SUBAPPLICATION Uebung_OPC_L16b_AX (* Wie L16, aber: gelesen wird erst, wenn INCREMENTED die Berechnung gemeldet hat (statt direkt nach dem Schreiben) *)
  (* Standard: 61499-2; Description: Copyright (c) 2026 Meisterschulen am Ostbahnhof This program and the accompanying materials are made available under the terms of the Eclipse Public License 2.0 which is available at https://www.eclipse.org/legal/epl-2.0/ SPDX-License-Identifier: EPL-2.0 *)
  (* Version 1.0, 2026-10-18, Franz Höpfinger, Meisterschulen am Ostbahnhof, B-Version von L16: Lesen erst nach INCREMENTED.CNF *)
  PACKAGE Meins::OPC_UA_Lokal;
  IMPORT Meins::OPC_UA_Lokal::const::OpcUaLokal::L16B_INC_READ;
  IMPORT Meins::OPC_UA_Lokal::const::OpcUaLokal::L16B_INCD_WRITE;
  IMPORT Meins::OPC_UA_Lokal::const::OpcUaLokal::L16B_INC_CLIENT_WRITE;
  IMPORT Meins::OPC_UA_Lokal::const::OpcUaLokal::L16B_INCD_CLIENT_READ;
  IMPORT logiBUS::io::DI::logiBUS_DI::Input_I1;
  IMPORT logiBUS::io::DI::logiBUS_DI_Events::BUTTON_PRESS_DOWN;
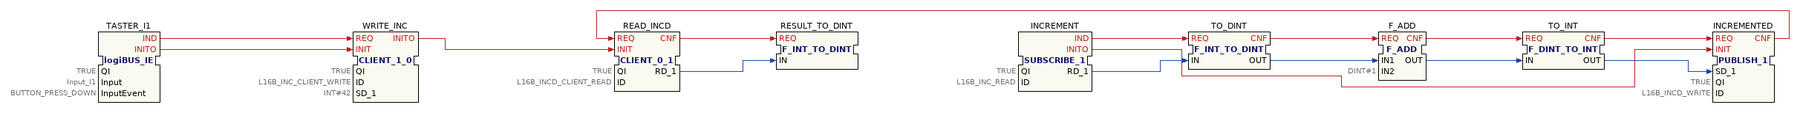
  (* B-Version von Uebung_OPC_L16_AX: READ_INCD.REQ kommt von INCREMENTED.CNF (Ergebnis ist veroeffentlicht), nicht von WRITE_INC.CNF. Das Lesen haengt so nicht mehr von der Reihenfolge ab. *)
  FBS
    TASTER_I1 : logiBUS::io::DI::logiBUS_IE(QI := TRUE, Input := Input_I1, InputEvent := BUTTON_PRESS_DOWN);
    WRITE_INC : iec61499::net::CLIENT_1_0(QI := TRUE, ID := L16B_INC_CLIENT_WRITE, SD_1 := INT#42);
    READ_INCD : iec61499::net::CLIENT_0_1(QI := TRUE, ID := L16B_INCD_CLIENT_READ);
    RESULT_TO_DINT : iec61131::conversion::F_INT_TO_DINT;
    INCREMENT : iec61499::net::SUBSCRIBE_1(QI := TRUE, ID := L16B_INC_READ);
    TO_DINT : iec61131::conversion::F_INT_TO_DINT;
    F_ADD : iec61131::arithmetic::F_ADD(IN2 := DINT#1);
    TO_INT : iec61131::conversion::F_DINT_TO_INT;
    INCREMENTED : iec61499::net::PUBLISH_1(QI := TRUE, ID := L16B_INCD_WRITE);
  END_FBS
  EVENT_CONNECTIONS
    TASTER_I1.IND TO WRITE_INC.REQ;
    INCREMENTED.CNF TO READ_INCD.REQ;
    TASTER_I1.INITO TO WRITE_INC.INIT;
    WRITE_INC.INITO TO READ_INCD.INIT;
    READ_INCD.CNF TO RESULT_TO_DINT.REQ;
    INCREMENT.IND TO TO_DINT.REQ;
    TO_DINT.CNF TO F_ADD.REQ;
    F_ADD.CNF TO TO_INT.REQ;
    TO_INT.CNF TO INCREMENTED.REQ;
    INCREMENT.INITO TO INCREMENTED.INIT;
  END_CONNECTIONS
  DATA_CONNECTIONS
    READ_INCD.RD_1 TO RESULT_TO_DINT.IN;
    INCREMENT.RD_1 TO TO_DINT.IN;
    TO_DINT.OUT TO F_ADD.IN1;
    F_ADD.OUT TO TO_INT.IN;
    TO_INT.OUT TO INCREMENTED.SD_1;
  END_CONNECTIONS
END_SUBAPPLICATION
